Fanuc KAREL source: kx00015.KL

-- PROVISIONAL review KL for V1013-1; original PC SHA256 9fa92da0ceaebeb69b251c188f9fcfea48370d380a0acb0726a4adbad6b07d60
-- Incomplete behavior may be omitted. Consult companion uncertainty JSON. Do not deploy.
PROGRAM KX00015
%NOLOCKGROUP
VAR
  I : INTEGER
  J : INTEGER
  B : BOOLEAN
  F : FILE
  S : STRING[80]
-- UNRESOLVED_DECL P type=000102
BEGIN
  -- UNRESOLVED_PC offsets 5-7; opcodes 9D,0E
  -- UNRESOLVED_PC offsets 12-16; opcodes 7F
END KX00015
